(* 소형 케이스 조립·검사·포장 자동화 공정 설계 *)

PROGRAM main
  VAR
    StartPB AT %IX0.0 : BOOL; (* 운전 시작 *)
    StopPB AT %IX0.1 : BOOL; (* 운전 정지 *)
    BodyDetected AT %IX0.2 : BOOL; (* 본체 투입 감지 *)
    LidDetected AT %IX0.3 : BOOL; (* 뚜껑 투입 감지 *)
    BodyAtAssembly AT %IX0.4 : BOOL; (* 본체 조립 위치 도착 *)
    LidAtAssembly AT %IX0.5 : BOOL; (* 뚜껑 조립 위치 도착 *)
    RobotReady AT %IX0.6 : BOOL; (* 로봇 작업 가능 *)
    RobotDone AT %IX0.7 : BOOL; (* 로봇 작업 완료 *)
    AssembledDetected AT %IX1.0 : BOOL; (* 조립품 배출 감지 *)
    InspectionDetected AT %IX1.1 : BOOL; (* 검사 위치 도착 *)
    RejectDetected AT %IX1.2 : BOOL; (* 불량품 배출 확인 *)
    PackDetected AT %IX1.3 : BOOL; (* 포장 위치 도착 *)
    PackDone AT %IX1.4 : BOOL; (* 포장 완료 *)
    FinishedGoodsDetected AT %IX1.5 : BOOL; (* 완제품 이동 확인 *)
    ShipmentDetected AT %IX1.6 : BOOL;
    SortEye AT %IX2.2 : BOOL; (* 불량 분기 위치 감지 *)
    PackDonePulse : BOOL;
    BodyLaunchPulse : BOOL;
    RejectPulse : BOOL;
    ShipPulse : BOOL;
    FeedPermit : BOOL;
    TargetShipped : BOOL;
    LaunchAllowance : UINT;
    LaunchedCount AT %MW111 : UINT;
    ShippedCount AT %MW110 : UINT;
    M16 : BOOL; (* 조립품 배출 시 한 번만 다음 사이클 허가 *)
    AssemblyJoinedSim AT %IX2.4 : BOOL; (* OIP 조립품 결합 완료 *)
    RobotReleasedSignal AT %QX2.0 : BOOL; (* OIP 조립 셀에 로봇 완료 전달 *) (* 출고 위치 통과 확인 *)
    BodyConveyorRun AT %QX0.0 : BOOL; (* 본체 컨베이어 가동 *)
    LidConveyorRun AT %QX0.1 : BOOL; (* 뚜껑 컨베이어 가동 *)
    BodyFeedEnable AT %QX0.2 : BOOL; (* 본체 공급 허가 *)
    LidFeedEnable AT %QX0.3 : BOOL; (* 뚜껑 공급 허가 *)
    BodyStopper AT %QX0.4 : BOOL; (* 본체 정위치 정지 *)
    LidStopper AT %QX0.5 : BOOL; (* 뚜껑 정위치 정지 *)
    RobotStart AT %QX0.6 : BOOL; (* 로봇 작업 시작 *)
    AssemblyOutRun AT %QX0.7 : BOOL; (* 조립품 배출 *)
    InspectionConveyorRun AT %QX1.0 : BOOL; (* 검사 컨베이어 가동 *)
    RejectDiverter AT %QX1.1 : BOOL; (* 불량품 분기 *)
    PackingConveyorRun AT %QX1.2 : BOOL; (* 포장 컨베이어 가동 *)
    PackStart AT %QX1.3 : BOOL; (* 포장 작업 시작 *)
    FinishedGoodsConveyorRun AT %QX1.4 : BOOL; (* 완제품 이송 *)
    ShippingConveyorRun AT %QX1.5 : BOOL; (* 출고 컨베이어 가동 *)
    AlarmLamp AT %QX1.6 : BOOL; (* 설비 이상 표시 *)
    WorkOrderActive AT %MW100 : UINT; (* 생산지시 활성화 (0/1) *)
    ProductType AT %MW101 : UINT; (* 제품 종류 번호 *)
    TargetQuantity AT %MW102 : UINT; (* 생산 목표 수량 *)
    MaterialPermit AT %MW103 : UINT; (* 자재 공급 허가 (0/1) *)
    ProducedCount AT %MW104 : UINT; (* 누적 생산 완료 수량 *)
    RejectCount AT %MW105 : UINT; (* 누적 불량 수량 *)
    MachineState AT %MW106 : UINT; (* 설비 운전 상태 코드  0 - IDLE : 생산 대기 1 - READY : 운전 준비 완료 2 - RUNNING : 생산 중 3 - MATERIAL_WAIT : 자재 부족 대기 4 - STOPPED : 정상 정지 5 - FAULT : 설비 오류 6 - COMPLETE : 생산 목표 완료 *)
    FaultCode AT %MW107 : UINT; (* 오류 원인 코드 *)
    InspectionResultValidWord AT %MW108 : UINT; (* 품질 검사 완료 여부(0/1) *)
    InspectionResultValid : BOOL; (* 품질 검사 완료 여부(0/1) => boolean 값으로 변환 *)
    InspectionResultWord AT %MW109 : UINT; (* 품질 검사 결과(0/1) *)
    InspectionResult : BOOL; (* 품질 검사 결과(0/1) => boolean 값으로 변환 *)
    WorkOrderActiveOK : BOOL; (* 생산지시 활성화 (0/1) => boolean 값으로 변환 *)
    M0 : BOOL; (* 생산 허가 : 운전 가동 릴레이 : M0 *)
    M1 : BOOL; (* 본체 투입 감지 릴레이 *)
    M2 : BOOL; (* 뚜껑 투입 감지 릴레이 *)
    M3 : BOOL; (* 본체 조립 위치 도착 릴레이 *)
    M4 : BOOL; (* 뚜껑 조립 위치 도착 릴레이 *)
    M5 : BOOL; (* 로봇 작업 가능 릴레이 *)
    M6 : BOOL; (* 로봇 작업 완료 릴레이 *)
    M7 : BOOL; (* 조립품 배출 감지 릴레이 *)
    M8 : BOOL; (* 검사 위치 도착 릴레이 *)
    M9 : BOOL; (* 품질 검사 완료 릴레이 *)
    M10 : BOOL; (* 품질 검사 결과가 불량품일 경우 불량품 배출 감지 릴레이 *)
    M11 : BOOL; (* 품질 검사 결과가 온품인 릴레이 *)
    M12 : BOOL; (* 포장 위치 도착 릴레이 *)
    M13 : BOOL; (* 포장 완료 릴레이 *)
    M14 : BOOL; (* 완제품 이송 감지 릴레이 *)
    M15 : BOOL; (* 출고 위치 통과 감지 릴레이 *)
  END_VAR

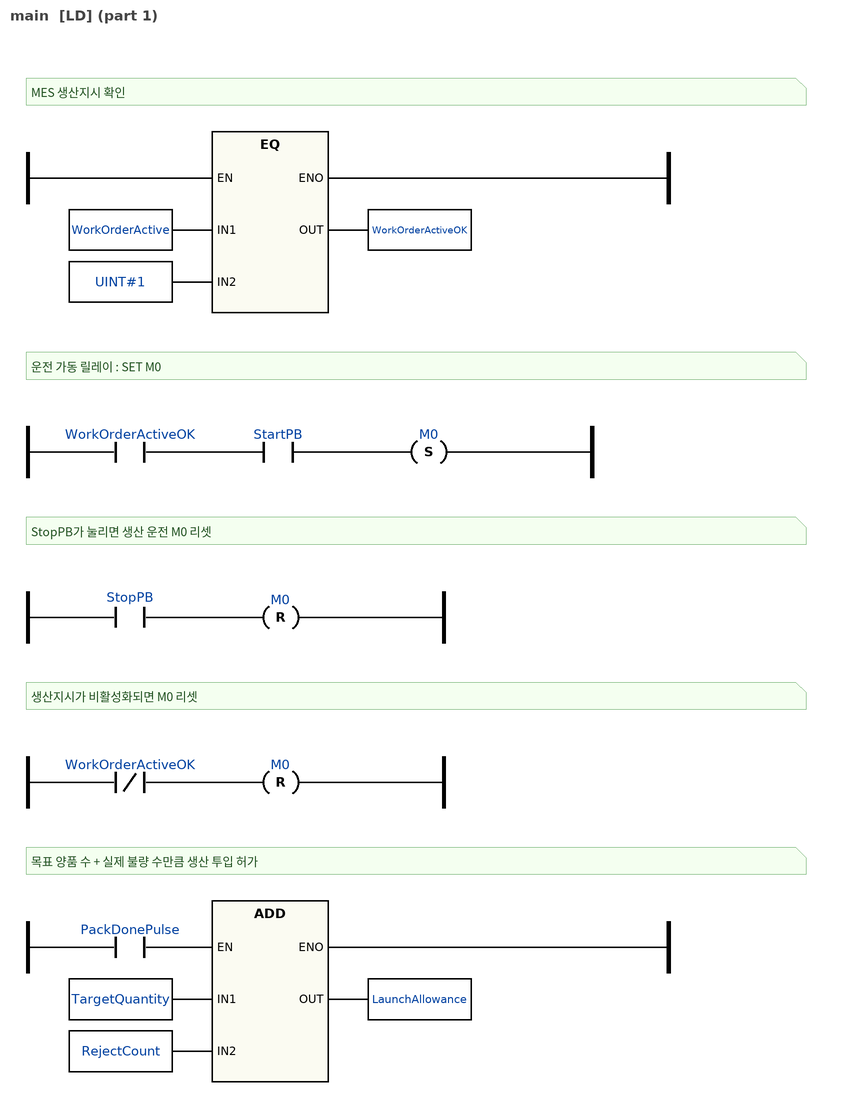
(* LD diagram, written out as Structured Text *)
(* MES 생산지시 확인 *)
WorkOrderActiveOK := WorkOrderActive = UINT#1;
(* 운전 가동 릴레이 : SET M0 *)
IF WorkOrderActiveOK AND StartPB THEN M0 := TRUE; END_IF;
(* StopPB가 눌리면 생산 운전 M0 리셋 *)
IF StopPB THEN M0 := FALSE; END_IF;
(* 생산지시가 비활성화되면 M0 리셋 *)
IF NOT WorkOrderActiveOK THEN M0 := FALSE; END_IF;
(* 목표 양품 수 + 실제 불량 수만큼 생산 투입 허가 *)
IF PackDonePulse THEN LaunchAllowance := TargetQuantity + RejectCount; END_IF;
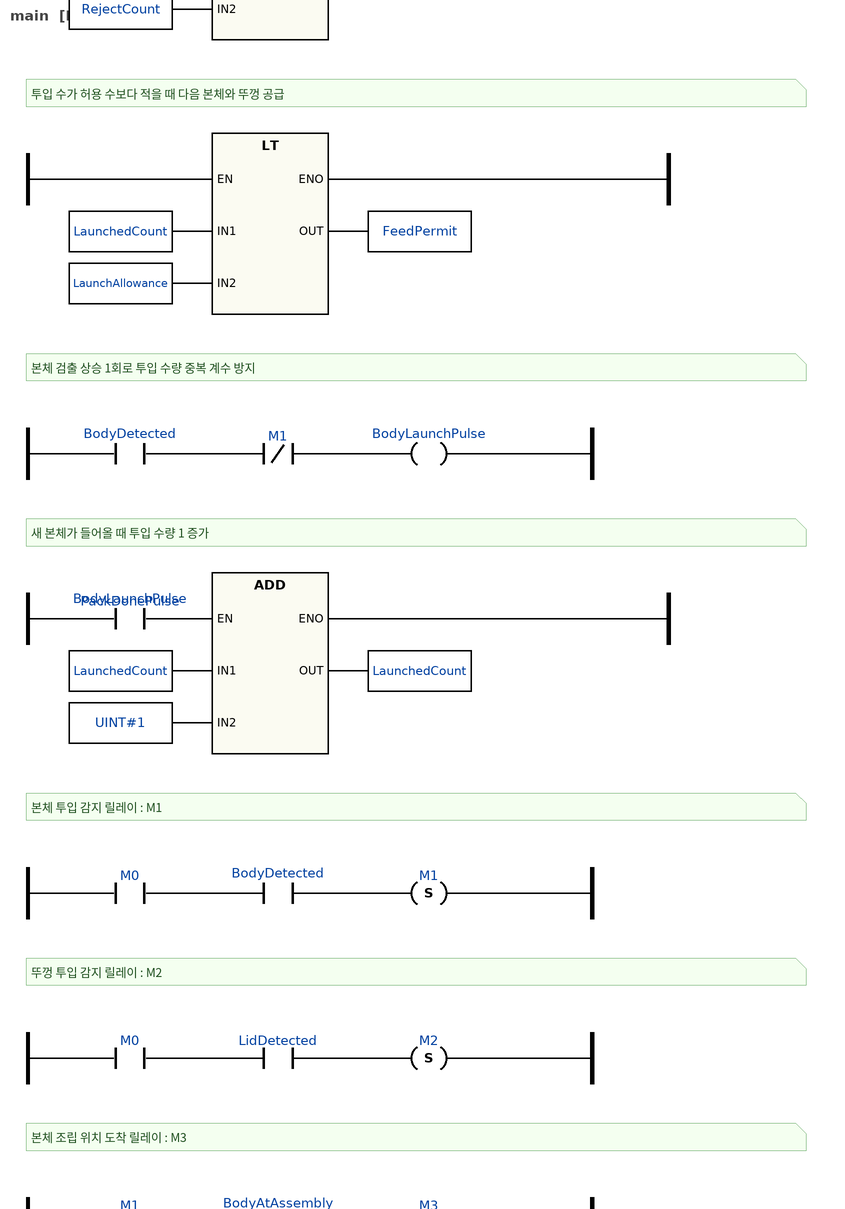
(* 투입 수가 허용 수보다 적을 때 다음 본체와 뚜껑 공급 *)
FeedPermit := LaunchedCount < LaunchAllowance;
(* 본체 검출 상승 1회로 투입 수량 중복 계수 방지 *)
BodyLaunchPulse := BodyDetected AND NOT M1;
(* 새 본체가 들어올 때 투입 수량 1 증가 *)
IF PackDonePulse AND BodyLaunchPulse THEN LaunchedCount := LaunchedCount + UINT#1; END_IF;
(* 본체 투입 감지 릴레이 : M1 *)
IF M0 AND BodyDetected THEN M1 := TRUE; END_IF;
(* 뚜껑 투입 감지 릴레이 : M2 *)
IF M0 AND LidDetected THEN M2 := TRUE; END_IF;
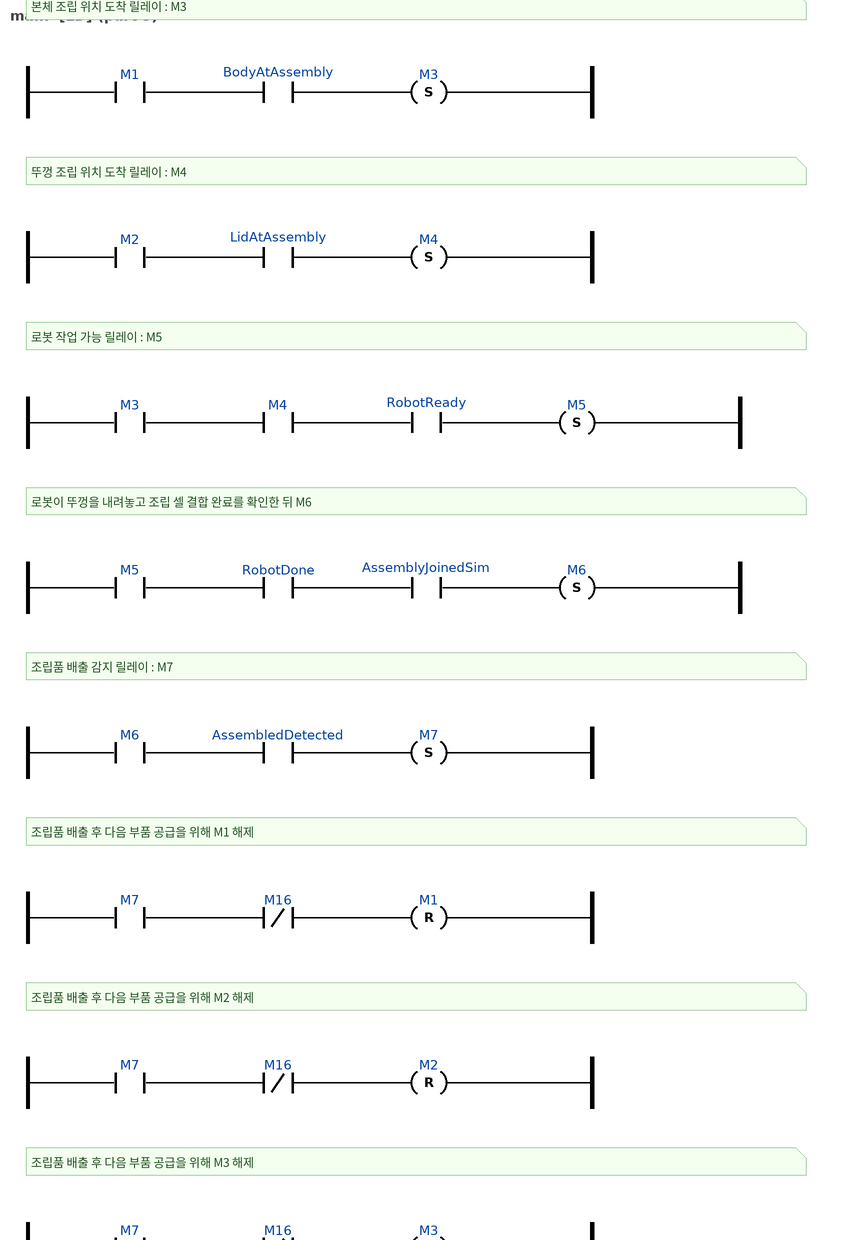
(* 본체 조립 위치 도착 릴레이 : M3 *)
IF M1 AND BodyAtAssembly THEN M3 := TRUE; END_IF;
(* 뚜껑 조립 위치 도착 릴레이 : M4 *)
IF M2 AND LidAtAssembly THEN M4 := TRUE; END_IF;
(* 로봇 작업 가능 릴레이 : M5 *)
IF M3 AND M4 AND RobotReady THEN M5 := TRUE; END_IF;
(* 로봇이 뚜껑을 내려놓고 조립 셀 결합 완료를 확인한 뒤 M6 *)
IF M5 AND RobotDone AND AssemblyJoinedSim THEN M6 := TRUE; END_IF;
(* 조립품 배출 감지 릴레이 : M7 *)
IF M6 AND AssembledDetected THEN M7 := TRUE; END_IF;
(* 조립품 배출 후 다음 부품 공급을 위해 M1 해제 *)
IF M7 AND NOT M16 THEN M1 := FALSE; END_IF;
(* 조립품 배출 후 다음 부품 공급을 위해 M2 해제 *)
IF M7 AND NOT M16 THEN M2 := FALSE; END_IF;
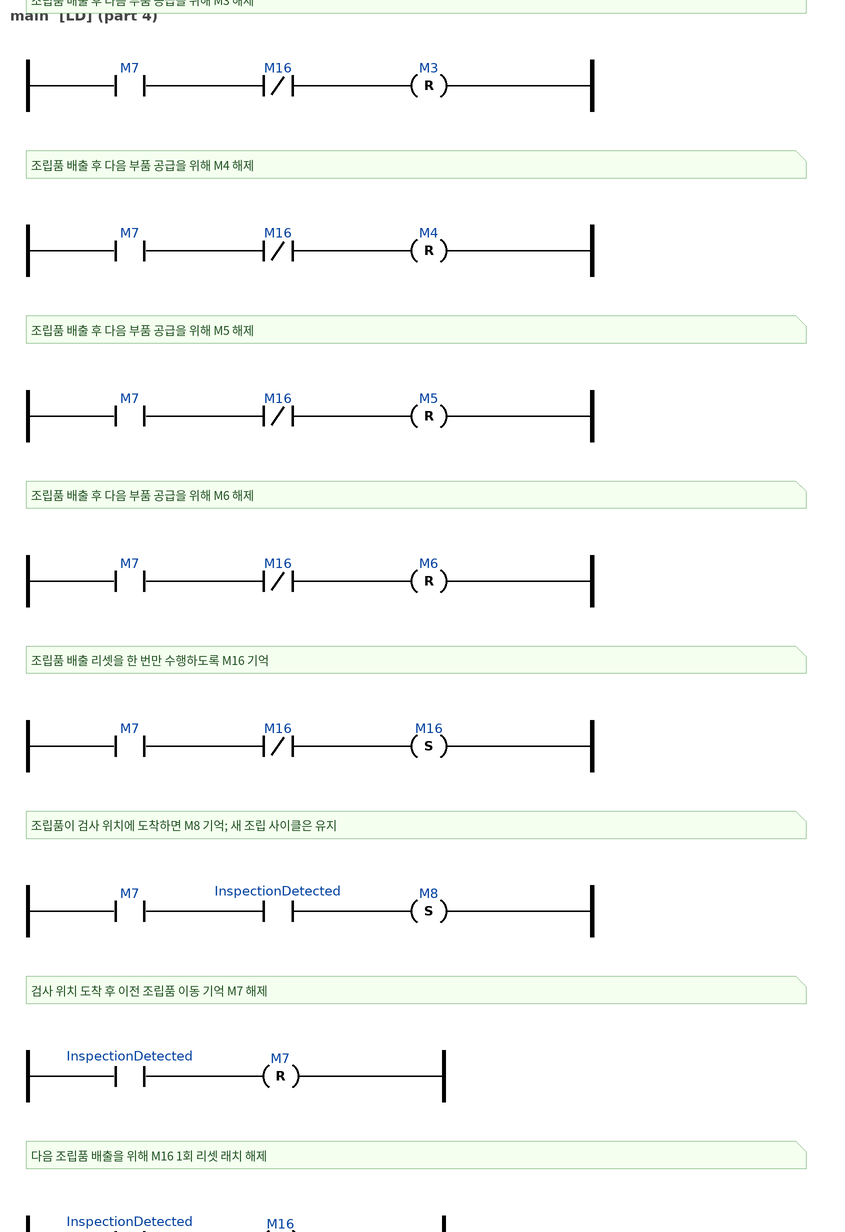
(* 조립품 배출 후 다음 부품 공급을 위해 M3 해제 *)
IF M7 AND NOT M16 THEN M3 := FALSE; END_IF;
(* 조립품 배출 후 다음 부품 공급을 위해 M4 해제 *)
IF M7 AND NOT M16 THEN M4 := FALSE; END_IF;
(* 조립품 배출 후 다음 부품 공급을 위해 M5 해제 *)
IF M7 AND NOT M16 THEN M5 := FALSE; END_IF;
(* 조립품 배출 후 다음 부품 공급을 위해 M6 해제 *)
IF M7 AND NOT M16 THEN M6 := FALSE; END_IF;
(* 조립품 배출 리셋을 한 번만 수행하도록 M16 기억 *)
IF M7 AND NOT M16 THEN M16 := TRUE; END_IF;
(* 조립품이 검사 위치에 도착하면 M8 기억; 새 조립 사이클은 유지 *)
IF M7 AND InspectionDetected THEN M8 := TRUE; END_IF;
(* 검사 위치 도착 후 이전 조립품 이동 기억 M7 해제 *)
IF InspectionDetected THEN M7 := FALSE; END_IF;
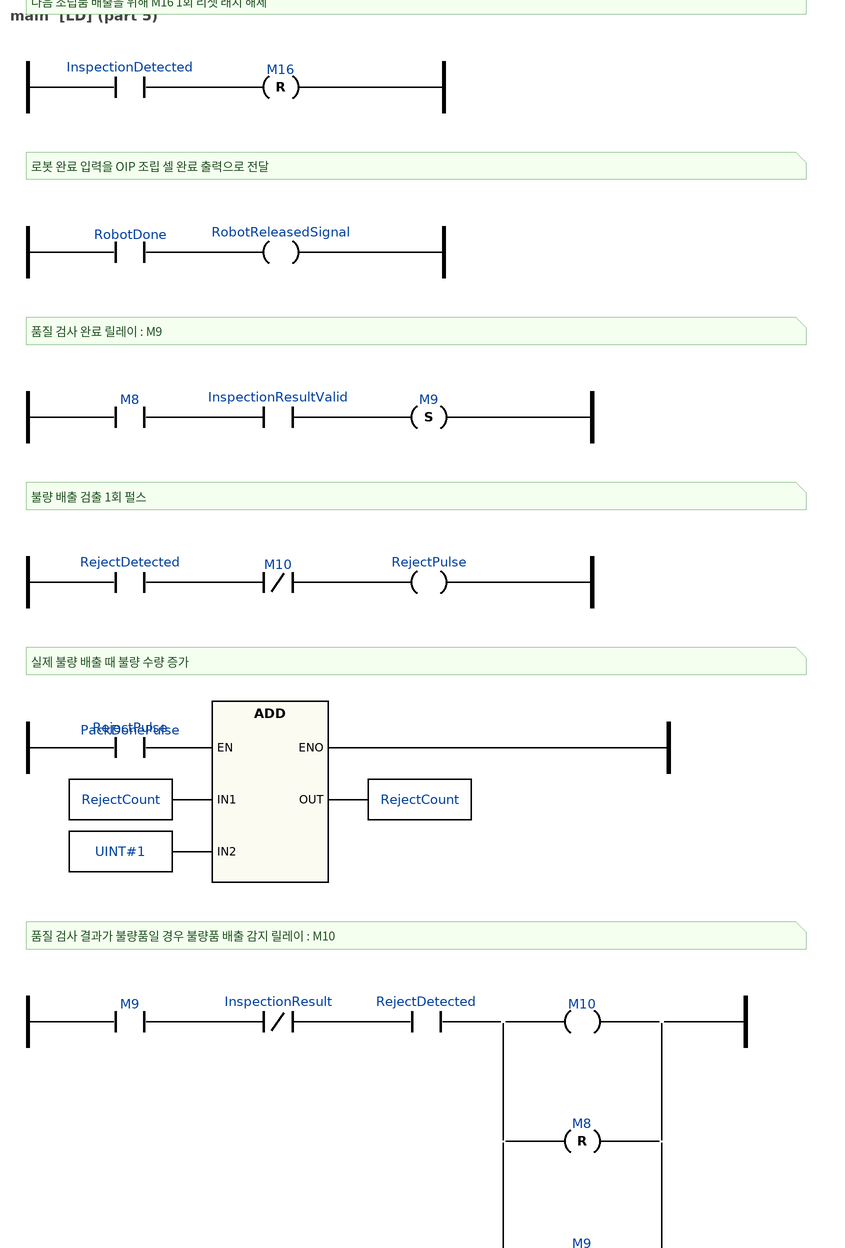
(* 다음 조립품 배출을 위해 M16 1회 리셋 래치 해제 *)
IF InspectionDetected THEN M16 := FALSE; END_IF;
(* 로봇 완료 입력을 OIP 조립 셀 완료 출력으로 전달 *)
RobotReleasedSignal := RobotDone;
(* 품질 검사 완료 릴레이 : M9 *)
IF M8 AND InspectionResultValid THEN M9 := TRUE; END_IF;
(* 불량 배출 검출 1회 펄스 *)
RejectPulse := RejectDetected AND NOT M10;
(* 실제 불량 배출 때 불량 수량 증가 *)
IF PackDonePulse AND RejectPulse THEN RejectCount := RejectCount + UINT#1; END_IF;
(* 품질 검사 결과가 불량품일 경우 불량품 배출 감지 릴레이 : M10 *)
M10 := M9 AND NOT InspectionResult AND RejectDetected;
IF M9 AND NOT InspectionResult AND RejectDetected THEN M8 := FALSE; END_IF;
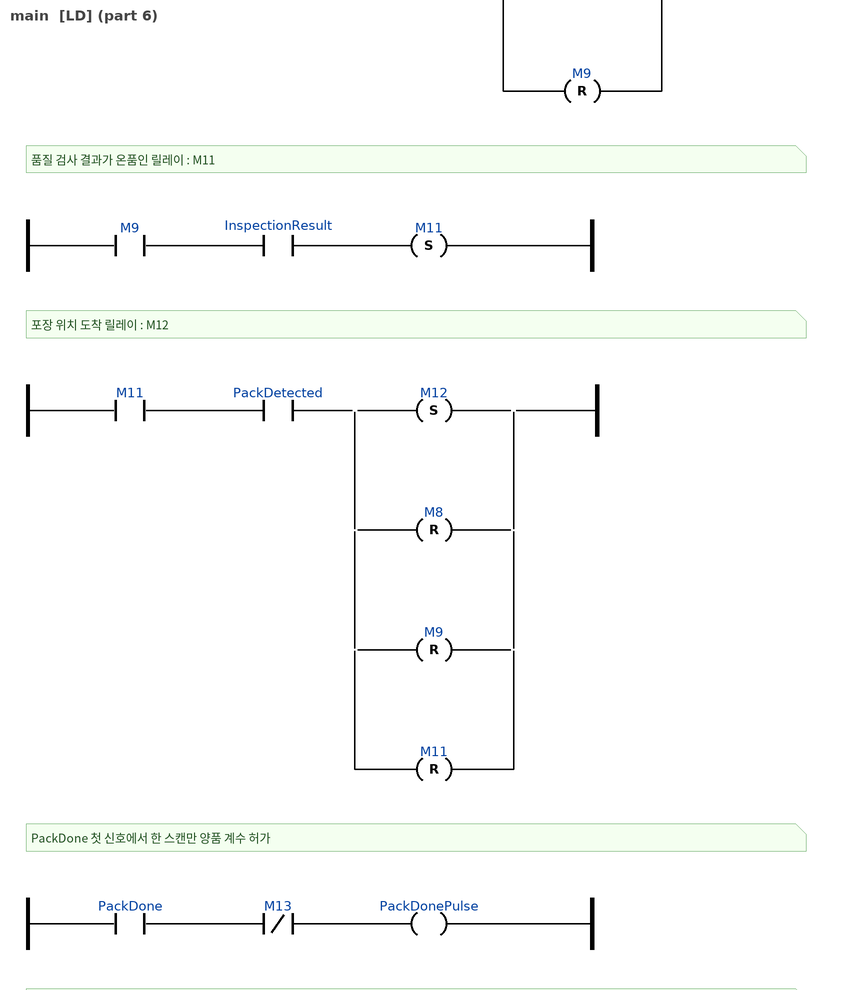
IF M9 AND NOT InspectionResult AND RejectDetected THEN M9 := FALSE; END_IF;
(* 품질 검사 결과가 온품인 릴레이 : M11 *)
IF M9 AND InspectionResult THEN M11 := TRUE; END_IF;
(* 포장 위치 도착 릴레이 : M12 *)
IF M11 AND PackDetected THEN M12 := TRUE; END_IF;
IF M11 AND PackDetected THEN M8 := FALSE; END_IF;
IF M11 AND PackDetected THEN M9 := FALSE; END_IF;
IF M11 AND PackDetected THEN M11 := FALSE; END_IF;
(* PackDone 첫 신호에서 한 스캔만 양품 계수 허가 *)
PackDonePulse := PackDone AND NOT M13;
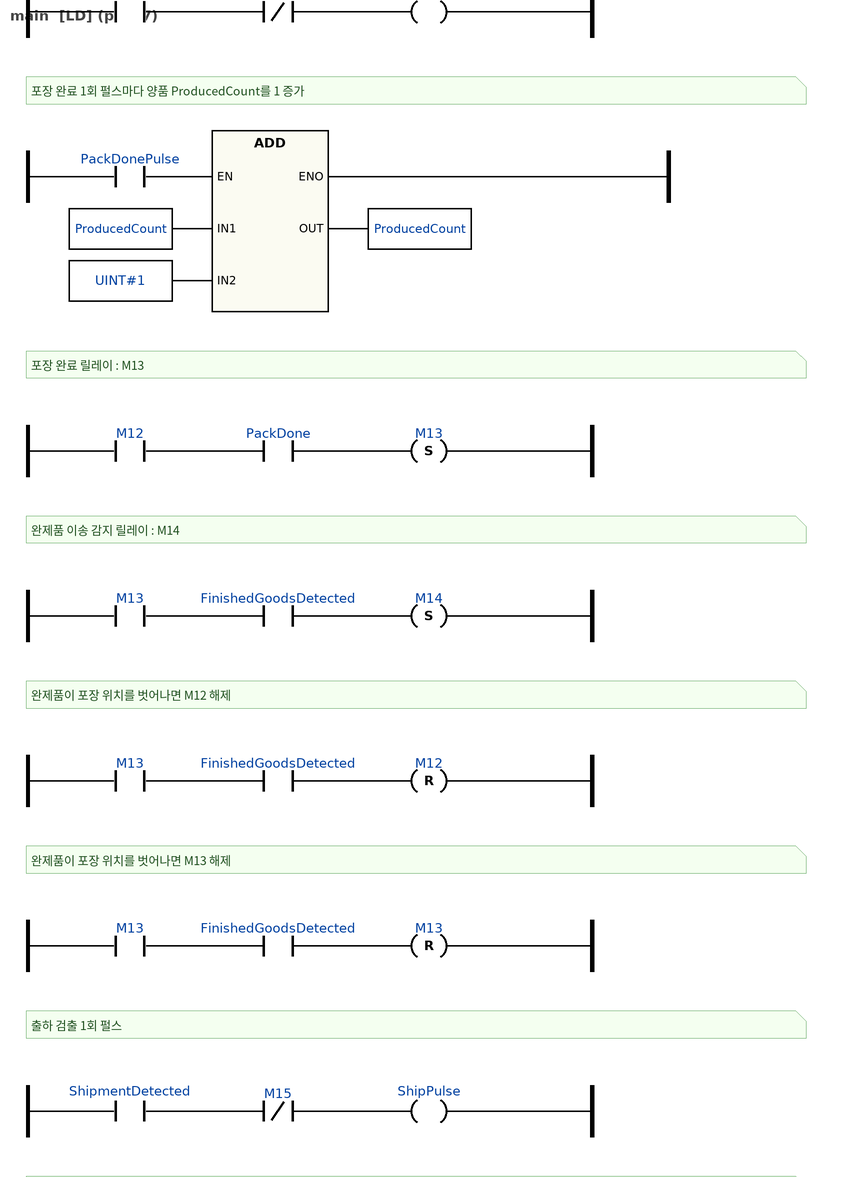
(* 포장 완료 1회 펄스마다 양품 ProducedCount를 1 증가 *)
IF PackDonePulse THEN ProducedCount := ProducedCount + UINT#1; END_IF;
(* 포장 완료 릴레이 : M13 *)
IF M12 AND PackDone THEN M13 := TRUE; END_IF;
(* 완제품 이송 감지 릴레이 : M14 *)
IF M13 AND FinishedGoodsDetected THEN M14 := TRUE; END_IF;
(* 완제품이 포장 위치를 벗어나면 M12 해제 *)
IF M13 AND FinishedGoodsDetected THEN M12 := FALSE; END_IF;
(* 완제품이 포장 위치를 벗어나면 M13 해제 *)
IF M13 AND FinishedGoodsDetected THEN M13 := FALSE; END_IF;
(* 출하 검출 1회 펄스 *)
ShipPulse := ShipmentDetected AND NOT M15;
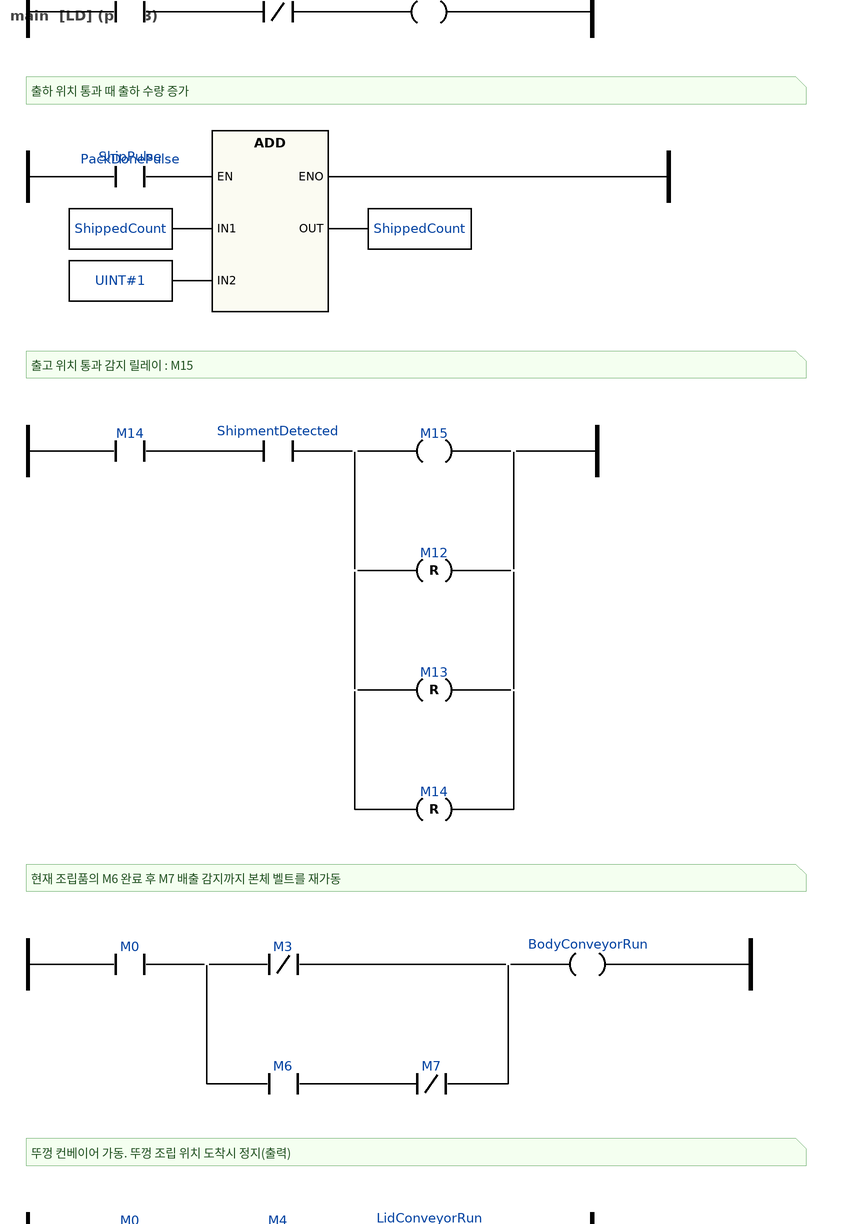
(* 출하 위치 통과 때 출하 수량 증가 *)
IF PackDonePulse AND ShipPulse THEN ShippedCount := ShippedCount + UINT#1; END_IF;
(* 출고 위치 통과 감지 릴레이 : M15 *)
M15 := M14 AND ShipmentDetected;
IF M14 AND ShipmentDetected THEN M12 := FALSE; END_IF;
IF M14 AND ShipmentDetected THEN M13 := FALSE; END_IF;
IF M14 AND ShipmentDetected THEN M14 := FALSE; END_IF;
(* 현재 조립품의 M6 완료 후 M7 배출 감지까지 본체 벨트를 재가동 *)
BodyConveyorRun := M0 AND (NOT M3 OR M6 AND NOT M7);
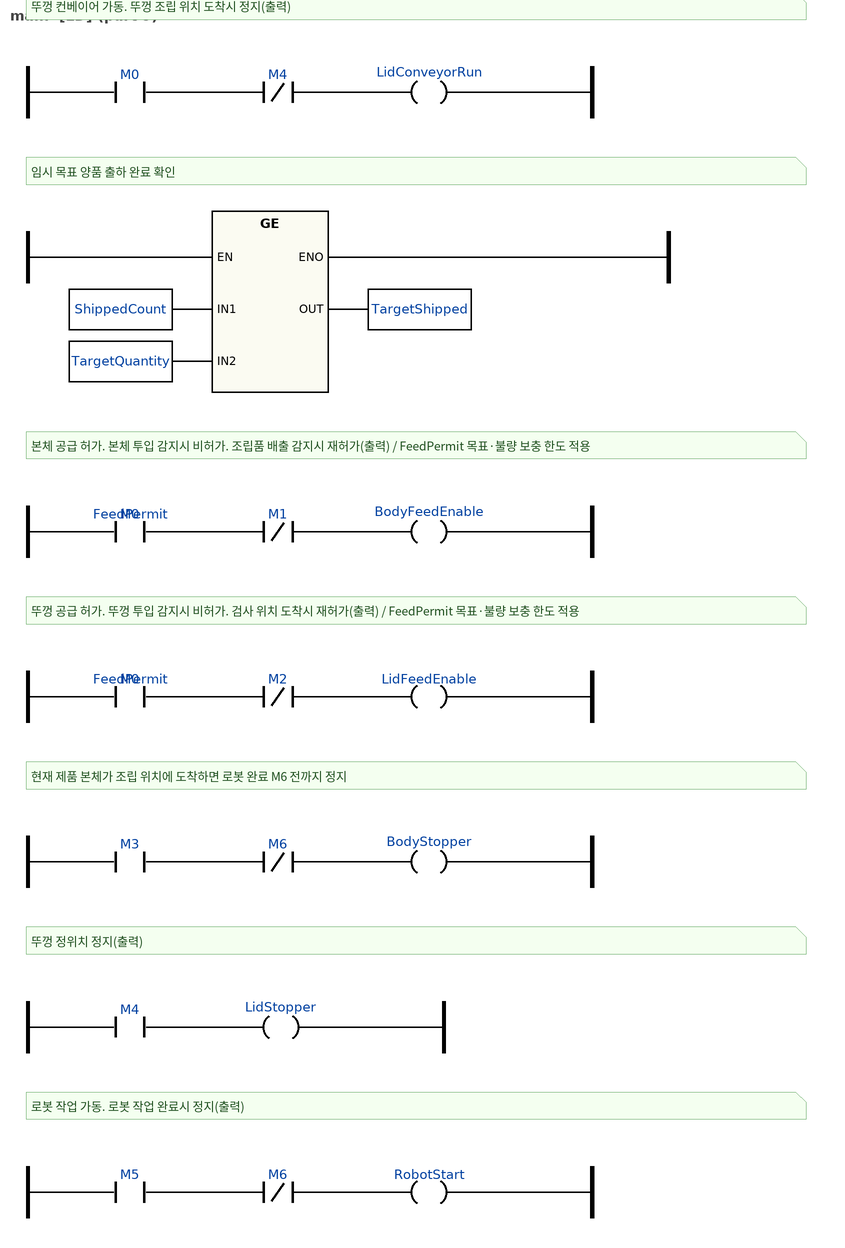
(* 뚜껑 컨베이어 가동. 뚜껑 조립 위치 도착시 정지(출력) *)
LidConveyorRun := M0 AND NOT M4;
(* 임시 목표 양품 출하 완료 확인 *)
TargetShipped := ShippedCount >= TargetQuantity;
(* 본체 공급 허가. 본체 투입 감지시 비허가. 조립품 배출 감지시 재허가(출력) / FeedPermit 목표·불량 보충 한도 적용 *)
BodyFeedEnable := M0 AND NOT M1 AND FeedPermit;
(* 뚜껑 공급 허가. 뚜껑 투입 감지시 비허가. 검사 위치 도착시 재허가(출력) / FeedPermit 목표·불량 보충 한도 적용 *)
LidFeedEnable := M0 AND NOT M2 AND FeedPermit;
(* 현재 제품 본체가 조립 위치에 도착하면 로봇 완료 M6 전까지 정지 *)
BodyStopper := M3 AND NOT M6;
(* 뚜껑 정위치 정지(출력) *)
LidStopper := M4;
(* 로봇 작업 가동. 로봇 작업 완료시 정지(출력) *)
RobotStart := M5 AND NOT M6;
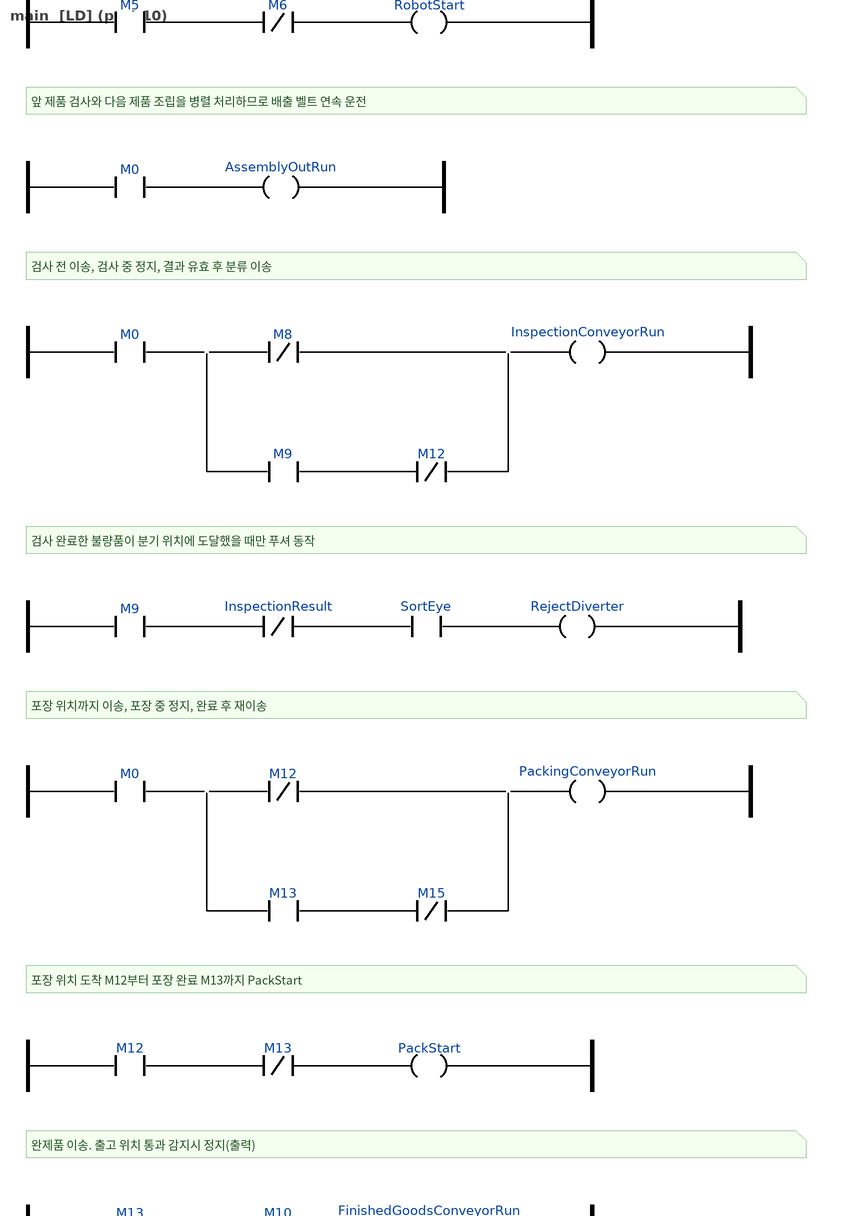
(* 앞 제품 검사와 다음 제품 조립을 병렬 처리하므로 배출 벨트 연속 운전 *)
AssemblyOutRun := M0;
(* 검사 전 이송, 검사 중 정지, 결과 유효 후 분류 이송 *)
InspectionConveyorRun := M0 AND (NOT M8 OR M9 AND NOT M12);
(* 검사 완료한 불량품이 분기 위치에 도달했을 때만 푸셔 동작 *)
RejectDiverter := M9 AND NOT InspectionResult AND SortEye;
(* 포장 위치까지 이송, 포장 중 정지, 완료 후 재이송 *)
PackingConveyorRun := M0 AND (NOT M12 OR M13 AND NOT M15);
(* 포장 위치 도착 M12부터 포장 완료 M13까지 PackStart *)
PackStart := M12 AND NOT M13;
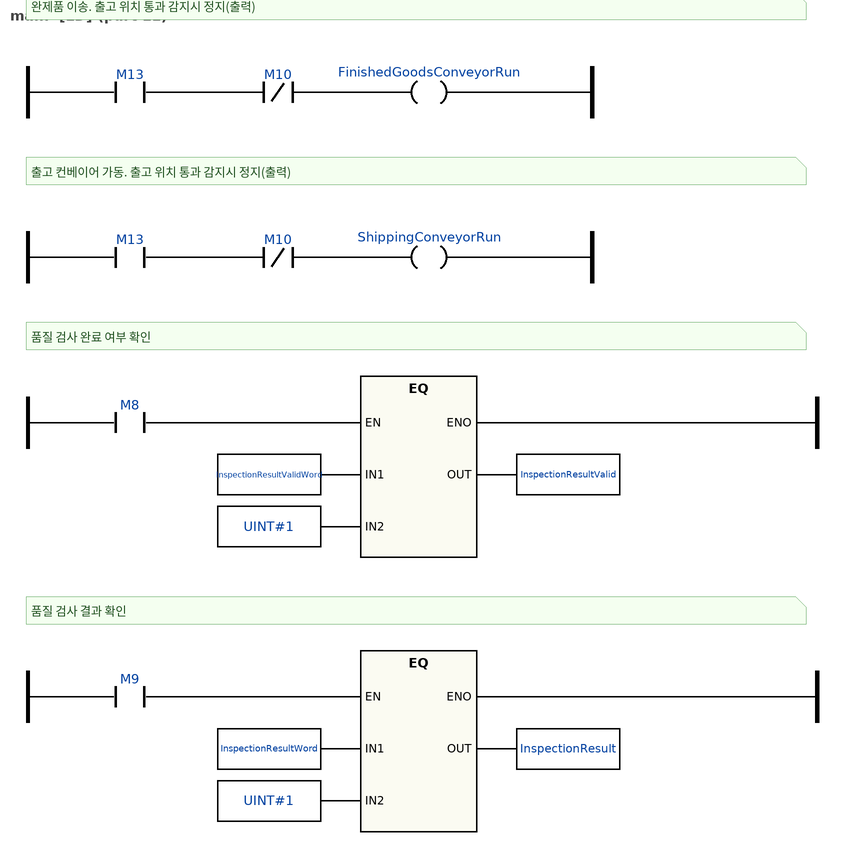
(* 완제품 이송. 출고 위치 통과 감지시 정지(출력) *)
FinishedGoodsConveyorRun := M13 AND NOT M10;
(* 출고 컨베이어 가동. 출고 위치 통과 감지시 정지(출력) *)
ShippingConveyorRun := M13 AND NOT M10;
(* 품질 검사 완료 여부 확인 *)
IF M8 THEN InspectionResultValid := InspectionResultValidWord = UINT#1; END_IF;
(* 품질 검사 결과 확인 *)
IF M9 THEN InspectionResult := InspectionResultWord = UINT#1; END_IF;
END_PROGRAM
